RoboDK station: вариант-1.rdk

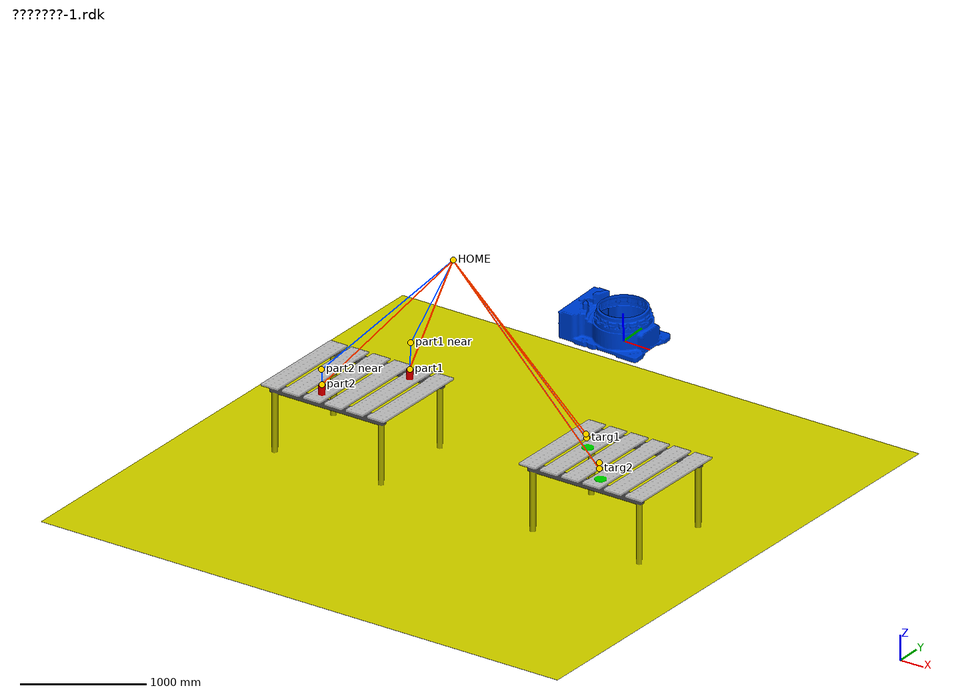
[picture v0: the station drawn from its stored meshes, robots at their saved joint values, targets as dots, program paths as lines]
Station вариант-1 (saved by RoboDK 6.0.6). Poses are relative to the parent item; angles as X-Y-Z fixed-axis rotations.
Station parameters (name, value as stored): LIN64
  - object Source table at (0, 0, 0) mm, size 1193.8 x 965.2 x 609.6 mm, geometry from welding_table.sld
  - object Destination table at (2500, 0, 0) mm, size 1193.8 x 965.2 x 609.6 mm, geometry from welding_table.sld
  - object Floor at (1190, 0, -610) mm, size 5000 x 5000 x 2.5 mm, geometry from plane_1m.sld
  - frame Yaskawa Motoman GP225 Base at (1499.86, 1544.03, 152.76) mm, rotated rx 2.47 ry 0.82 rz 0.04 deg
    - robot Yaskawa Motoman GP225: 6 axes, payload 225 kg, reach 3935 mm, repeatability 0.05 mm, weight 2702 kg
        joint limits [-180, -60, -86, -360, -125, -360] to [180, 76, 90, 360, 125, 360]; home [0, 0, 0, 0, 0, 0]; saved at [-100.341, -1.79, 1.132, -19.21, -8.061, 142.236]
      - tool OnRobot SG-b Soft Gripper, TCP at (0, 0, 150) mm, size 104 x 103.8 x 166.3 mm
    - target HOME (Cartesian target) at (-322.08, -1867.94, 1478.79) mm, rotated rx 95.59 ry 32.86 rz -4.65 deg; joints [-100.1, 5.55, 8.12, -18.37, -7.65, 141.4] of Yaskawa Motoman GP225
    - target part1 near (Cartesian target) at (-1179.48, -1260.38, 198.2) mm, rotated rx 177.39 ry -2.89 rz -40.49 deg; joints [-133.804, 11.973, -26.522, -4.014, -49.135, 95.815] of Yaskawa Motoman GP225
    - target part1 (Cartesian target) at (-1177.46, -1275.86, -31.27) mm, rotated rx 177.39 ry -2.89 rz -40.49 deg; joints [-133.398, 18.305, -30.489, -4.814, -38.844, 96.533] of Yaskawa Motoman GP225
    - target targ1 (Cartesian target) at (693.17, -1506.58, 12.47) mm, rotated rx 178.67 ry -2.59 rz 27.22 deg; joints [-65.934, 14.013, -33.669, -4.04, -41.201, 96.141] of Yaskawa Motoman GP225
    - target part2 near (Cartesian target) at (-1596.44, -1899.18, 122.5) mm, rotated rx 179.67 ry -1.73 rz -35.16 deg; joints [-130.332, 52.077, 29.906, -1.892, -67.668, 95.885] of Yaskawa Motoman GP225
    - target part2 (Cartesian target) at (-1593.56, -1902.16, -12.44) mm, rotated rx 179.67 ry -1.73 rz -35.16 deg; joints [-130.237, 53.815, 26.687, -1.969, -62.712, 95.974] of Yaskawa Motoman GP225
    - target targ2 (Cartesian target) at (1096.67, -1906.46, 40.76) mm, rotated rx -179.73 ry 1.8 rz 37.01 deg; joints [-59.76, 37.743, 2.16, 2.233, -54.497, 95.472] of Yaskawa Motoman GP225
    - target targ2 near (Cartesian target) at (1098.21, -1905.63, 95.73) mm, rotated rx -179.73 ry 1.8 rz 37.01 deg; joints [-59.715, 36.732, 3.224, 2.178, -56.572, 95.523] of Yaskawa Motoman GP225
    - target targ1 near (Cartesian target) at (691.39, -1506.58, 47.43) mm, rotated rx 178.67 ry -2.59 rz 27.22 deg; joints [-65.991, 12.971, -33.08, -3.916, -42.831, 96.029] of Yaskawa Motoman GP225
    - target Target 10 (Cartesian target) at (691.39, -1506.58, 47.43) mm, rotated rx 178.67 ry -2.59 rz 27.22 deg; joints [-65.991, 12.971, -33.08, -3.916, -42.831, 96.029] of Yaskawa Motoman GP225
    - target Target 11 (Cartesian target) at (691.39, -1506.58, 47.43) mm, rotated rx 178.67 ry -2.59 rz 27.22 deg; joints [-65.991, 12.971, -33.08, -3.916, -42.831, 96.029] of Yaskawa Motoman GP225
    - target Target 12 (Cartesian target) at (-322.08, -1867.94, 1478.79) mm, rotated rx 95.59 ry 32.86 rz -4.65 deg; joints [-100.341, -1.79, 1.132, -19.21, -8.061, 142.236] of Yaskawa Motoman GP225
  - program change (17 instructions, listed below)
  - object Target 1 at (2150, 0, 0) mm, size 100 x 99.9 x 10 mm, geometry from target.STL
  - program reset (16 instructions, listed below)
  - object Target 2 at (2560, -410, 0) mm, size 100 x 99.9 x 10 mm, geometry from target.STL
  - object Part 2 at (-90, -360, 40) mm, size 60 x 60 x 80 mm, geometry from part.sld
  - object Part 1 at (320, 270, 40) mm, size 60 x 60 x 80 mm, geometry from part.sld
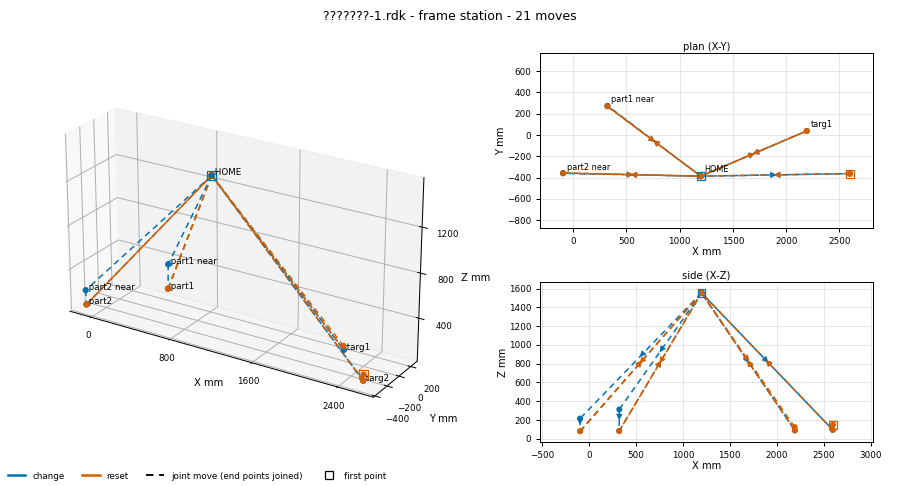
[picture p0: tool path of вариант-1.rdk in frame station, 21 of 21 moves have a stored position in this frame; points joined in program order, loops and branches not executed]

--- program change (robot Yaskawa Motoman GP225) ---
  Set Ref.: Yaskawa Motoman GP225 Base
  Set Tool: OnRobot SG-b Soft Gripper
  MoveJ (HOME)
  MoveJ (part1 near)
  MoveJ (part1)
  Attach to OnRobot SG-b Soft Gripper
  MoveJ (HOME)
  MoveJ (targ1)
  Detach from OnRobot SG-b Soft Gripper
  MoveJ (HOME)
  MoveJ (part2 near)
  MoveJ (part2)
  Attach to OnRobot SG-b Soft Gripper
  MoveJ (HOME)
  MoveJ (targ2)
  Detach from OnRobot SG-b Soft Gripper
  MoveJ (HOME)

--- program reset (robot Yaskawa Motoman GP225) ---
  Set Ref.: Yaskawa Motoman GP225 Base
  Set Tool: OnRobot SG-b Soft Gripper
  MoveJ (targ2 near)
  MoveJ (targ2)
  Attach to OnRobot SG-b Soft Gripper
  MoveJ (HOME)
  MoveJ (part2)
  Detach from OnRobot SG-b Soft Gripper
  MoveJ (HOME)
  MoveJ (targ1 near)
  MoveJ (targ1)
  Attach to OnRobot SG-b Soft Gripper
  MoveJ (HOME)
  MoveJ (part1)
  Detach from OnRobot SG-b Soft Gripper
  MoveJ (HOME)
